// TIA Portal V20 export
// export: Created 2026-10-20T12:41:04.2256983Z, ExportSetting WithDefaults, DisplayName Totally Integrated Automation Portal, DisplayVersion V20 Update 6, DisplayName TIA Portal Openness, DisplayVersion V20 Update 6, DisplayName TIA Portal Version Control Interface, DisplayVersion V20 Update 6, DisplayName SINAMICS Startdrive Advanced, DisplayVersion V20 SP1, DisplayName SINAMICS Startdrive G130, G150, S120, S150, SINAMICS MV, G220, S200, S210, DisplayVersion V20 SP1, DisplayName SINAMICS Startdrive G110M, G120, G120C, G120D, G120P, G115D, DisplayVersion V20 SP1, DisplayName STEP 7 Professional, DisplayVersion V20 Update 6, DisplayName STEP 7 Safety, DisplayVersion V20 Update 2, DisplayName WinCC Basic/Comfort/Advanced, DisplayVersion V20 Update 6, DisplayName WinCC Unified, DisplayVersion V20 Update 6
FUNCTION_BLOCK "SICK_Lector_Control_FB"   // FB19, SCL
{ S7_Optimized_Access := 'TRUE' }
VERSION : 0.1
// stored: AutoNumber true, IsIECCheckEnabled false, IsRetainMemResEnabled false, MemoryReserve 100, SetENOAutomatically false, UDAEnableTagReadback false
   VAR_INPUT
      Rd_Done : Bool;
      Req_Done : Bool;
      Req_Busy : Bool;
      Error : Bool;
      arrResult : Array[1..200] of Byte;
      iCounter : USInt;
      iLength : Int;
      Error_Code : DWord;
   END_VAR
   VAR_OUTPUT
      Test_Comm : Bool;
      Enable_Trigger : Bool;
      Disable_Trigger : Bool;
      Enable_Req : Bool;
      Result : String;
      Test_OK : Bool;
   END_VAR
   VAR_IN_OUT
      Test_Comm_HMI : Bool;
      Enable_HMI : Bool;
      Disable_HMI : Bool;
      Auto_Start_Lector : Bool;
      Auto_Stop_Lector : Bool;
   END_VAR
   VAR
      "Timer" { S7_SetPoint := 'True'} : TON_TIME;
      R_Done_DB { S7_SetPoint := 'True'} : R_TRIG;
      T_Reset_DB { S7_SetPoint := 'True'} : TON_TIME;
   END_VAR
BEGIN
   //Communication Test
   IF #Test_Comm_HMI THEN
       #Test_Comm := 1;
       #Enable_Req := 1;
       #Timer.TON(IN:=True,
                              PT:=t#1s);
   END_IF;

   //TEST OK
   IF #Req_Done AND #Timer.Q AND NOT #Error THEN
       #Test_OK := 1;
       #Test_Comm := 0;
       #Enable_Req := 0;
       #Test_Comm_HMI := 0;
       #Timer.TON(IN := FALSE,
                              PT := t#0s);
   END_IF;

   //ERROR
   IF #Timer.Q AND #Error THEN
           #Test_OK := 0;
           #Test_Comm := 0;
           #Enable_Req := 0;
           #Test_Comm_HMI := 0;
           #Timer.TON(IN := FALSE,
                                  PT := t#0s);
       END_IF;

   //Enable Trigger
       IF #Enable_HMI OR #Auto_Start_Lector THEN
       #Enable_Trigger := 1;
       #Enable_Req := 1;
       #Disable_HMI := 0;
       #Disable_Trigger := 0;
   //Disable Trigger
   ELSIF #Disable_HMI OR #"Auto_Stop_Lector" THEN
       #Disable_Trigger := 1;
       #Enable_Req := 1;
       #Enable_HMI := 0;
       #Enable_Trigger := 0;
   ELSE
       #Enable_Trigger := 0;
       #Enable_Req := 0;
       #Disable_Trigger := 0;
   END_IF;


   #R_Done_DB(CLK:=#Rd_Done);

   IF #R_Done_DB.Q OR #T_Reset_DB.Q OR
       (#Enable_HMI AND #Disable_HMI)
   THEN
       #Disable_HMI := 0;
       #Enable_Trigger := 0;
       #Disable_Trigger := 0;
       #Enable_Req := 0;
       #T_Reset_DB.TON(IN := FALSE,
                               PT := T#0S);
               #Auto_Stop_Lector := 0;
   END_IF;

   #T_Reset_DB(IN:=(#Enable_HMI OR #Disable_HMI OR #Auto_Start_Lector OR #Auto_Stop_Lector),
                 PT:=T#10S);


   #Result := "ByteArrayToString_1"(Lenght := #iLength, ByteArray := #arrResult);
END_FUNCTION_BLOCK
